(* IEC 61131-3 sources: codesys/project-view/Device/Plc Logic/Application/000-模组/本项目, 8 files *)

(* ---- FC_ArrayBoolHasTrue.st ---- *)
//布尔数组里面至少有一个值为true的话，函数返回TRUE
FUNCTION FC_ArrayBoolHasTrue : BOOL
VAR_IN_OUT
	abArray							: ARRAY[*] OF BOOL;
END_VAR

VAR
	i								: DINT;
END_VAR
// --- implementation ---
FOR i := LOWER_BOUND(abArray,1) TO UPPER_BOUND(abArray,1) DO
	IF abArray[i] THEN
		FC_ArrayBoolHasTrue := TRUE;
		RETURN;
	END_IF
END_FOR

FC_ArrayBoolHasTrue := FALSE;
END_FUNCTION

(* ---- FC_IsInArea.st ---- *)
FUNCTION FC_IsInArea : BOOL
VAR_INPUT
	LR_Pos							: REAL;//当前左右位置
	UD_Pos							: REAL;//当前上下位置

	LeftLimit						: REAL;//左边限位，LR_Pos要大于等于此变量
	RightLimit						: REAL;//右边限位，LR_Pos要小于等于此变量
	UpLimit							: REAL;//上边限位，UD_Pos要小于等于此变量
	DownLimit						: REAL;//下边限位，UD_Pos要大于等于此变量
END_VAR
VAR
END_VAR
// --- implementation ---
//判断是否在此平面范围内

IF (LeftLimit <= LR_Pos AND LR_Pos <= RightLimit) AND
	(DownLimit <= UD_Pos AND UD_Pos <= UpLimit) THEN

	FC_IsInArea := TRUE;
ELSE
	FC_IsInArea := FALSE;
END_IF
END_FUNCTION

(* ---- FC_StringConnect.st ---- *)
//输出 STRING = sStr1 + sStr2 + sStr3 + sStr4 +sStr5
FUNCTION FC_StringConnect : STRING
VAR_INPUT
	sStr1						: STRING:='';
	sStr2						: STRING:='';
	sStr3						: STRING:='';
	sStr4						: STRING:='';
	sStr5						: STRING:='';

END_VAR

VAR
	temp						: STRING;

END_VAR
// --- implementation ---
//temp := sStr1;

// StrConcatW(pstFrom:=ADR(wsContent_2) , pstTo:=ADR(temp) , iBufferSize:=TO_INT(SIZEOF(temp)) );
// StrConcatW(pstFrom:=ADR(wsContent_3) , pstTo:=ADR(temp) , iBufferSize:=TO_INT(SIZEOF(temp)) );

temp := CONCAT(STR1:=sStr1 , STR2:=sStr2 );
temp := CONCAT(STR1:=temp , STR2:=sStr3 );
temp := CONCAT(STR1:=temp , STR2:=sStr4 );
temp := CONCAT(STR1:=temp , STR2:=sStr5 );

FC_StringConnect := temp;
END_FUNCTION

(* ---- FC_WordToReal.st ---- *)
FUNCTION FC_WordToReal : REAL
VAR_INPUT
	arrRegisters0 : WORD;
	arrRegisters1 : WORD;
END_VAR
VAR
	dwCombined: DWORD;              // 合并后的DWORD
    rResult: REAL;                  // 输出浮点数
    pReal: POINTER TO REAL;         // 类型转换指针
    bIsBigEndian: BOOL := TRUE;     // 字节序配置开关
END_VAR
// --- implementation ---
// 寄存器合并与转换逻辑
IF bIsBigEndian THEN
    dwCombined := SHL(WORD_TO_DWORD(arrRegisters0), 16) OR arrRegisters1;
ELSE
    dwCombined := SHL(WORD_TO_DWORD(arrRegisters0), 16) OR arrRegisters1;
END_IF

pReal := ADR(dwCombined);           // 获取内存地址
FC_WordToReal := pReal^;                  // 指针解引用
END_FUNCTION

(* ---- FB_DelayInvert.st ---- *)
//X维持设定的初始值，直到指定时间结束，取反。
//若中途取消动作，X保持设定的初始值。
FUNCTION_BLOCK FB_DelayInvert
VAR_IN_OUT
	X							: BOOL;
END_VAR

VAR_INPUT
	bStart						: BOOL;
	bStop						: BOOL;

	bInitValue					: BOOL;//初始值
	tDelay						: TIME:=T#1S;

END_VAR

VAR_OUTPUT
END_VAR

VAR
	timer						: TON;
	R_TRIG_Start				: R_TRIG;
	R_TRIG_Stop					: R_TRIG;

END_VAR
// --- implementation ---
//定时器FB块
timer();

//启动
R_TRIG_Start(CLK:=bStart);
IF R_TRIG_Start.Q THEN
	X := bInitValue;
	timer.PT := tDelay;
	timer.IN := TRUE;
	bStart := FALSE;
END_IF

//定时器计时中（触发动作），中途取消动作，X维持初始值
R_TRIG_Stop(CLK:=bStop);
IF R_TRIG_Stop.Q AND timer.IN THEN
	X := bInitValue;
	timer.IN := FALSE;
END_IF

//时间到，取反
IF timer.Q THEN
	X := NOT X;
	timer.IN := FALSE;
END_IF
END_FUNCTION_BLOCK

(* ---- FB_Overtime.st ---- *)
FUNCTION_BLOCK FB_Overtime
VAR_INPUT
	bEnable						: BOOL;
	tTimeSet					: TIME:=T#1S;//定时时间
	iMode						: INT:=0;//超时后，0模式的bEnable变false，输出跟着变false；1模式的bEnable变false，输出不变，需要bReset复位。
	bReset						: BOOL;//上升沿将输出复位为false，仅1模式有效
END_VAR

VAR_OUTPUT
	bOvertime					: BOOL;
END_VAR

VAR
	tTimer						: TON;
	R_TRIG_1						: R_TRIG;
	R_TRIG_2						: R_TRIG;
END_VAR
// --- implementation ---
tTimer(IN:=bEnable , PT:= tTimeSet);
R_TRIG_1(CLK:=tTimer.Q);
R_TRIG_2(CLK:=bReset);

IF iMode = 0 THEN
	IF tTimer.Q THEN
		bOvertime:=TRUE;
	ELSE
		bOvertime:=FALSE;
	END_IF

ELSIF iMode = 1 THEN
	IF R_TRIG_1.Q THEN
		bOvertime:=TRUE;
	END_IF
	IF R_TRIG_2.Q THEN
		bOvertime:=false;
	END_IF

END_IF
END_FUNCTION_BLOCK

(* ---- FB_TcpClient_Free_1.st ---- *)
FUNCTION_BLOCK FB_TcpClient_Free_1
VAR_INPUT
	xConnect			:BOOL;				//连接
	xDisConnect			:BOOL;				//断开连接
	xReset				:BOOL;				//复位
	strIP				:STRING;			//IP
	uiPort				:UINT;				//端口号
	xSend				:BOOL;				//发送
	pbySendData			:POINTER TO BYTE;	//发送数据变量容器起始地址
	uxiSendDataSize		:__UXINT;			//发送数据变量容器大小
	uxiSendLenght		:__UXINT;			//发送数据长度
	pbyReceiveData		:POINTER TO BYTE;	//接收数据变量容器起始地址
	uxiReceiveDataSize	:__UXINT;			//接收数据变量容器大小
END_VAR
VAR_OUTPUT
	xBusy				:BOOL;				//运行中
	xConnected			:BOOL;				//已连接
	xError				:BOOL;				//错误
	xSendDone			:BOOL;				//发送完毕
	udiNumOfSend		:UDINT;				//发送次数（满4294967295自动清零）
	xReceiveDone		:BOOL;				//接收完毕
	udiNumOfReceive		:UDINT;				//接收次数（满4294967295自动清零）
	udiReceiveLenght	:UDINT;				//接收数据长度
END_VAR
VAR
	iStep			:INT;
	udiIndex		:UDINT;;
	fbClient		:TCP.Connector;
	eClientError	:TCP.ERROR;
	rtrigSend		:Standard.R_TRIG;
	eSendError		:TCP.ERROR;
	rtrigReceive	:Standard.R_TRIG;
	eReceiveError	:TCP.ERROR;
	xiReceiveLen	:__XINT;
	pby1			:POINTER TO BYTE;
	ton1:		Standard.TON;
END_VAR
// --- implementation ---
// ton1(IN:= TRUE, PT:= T#5000MS, Q=> , ET=> );
// IF NOT ton1.Q THEN
// 	RETURN;
// END_IF

IF xDisConnect THEN
	iStep:=0;
END_IF

//work step
CASE iStep OF

0:	//start
	fbClient.Disconnect();
	fbClient.Reset();
	RESET();
	xBusy:=FALSE;
	IF xConnect AND NOT xDisConnect THEN
		START();
		xBusy:=TRUE;
		iStep:=10;
	END_IF

10:	//wait connect
	eClientError:=fbClient.Connect(sIPAddress:= strIP, uiPort:= uiPort, pStream=> );
	IF eClientError = TCP.ERROR.NO_ERROR THEN
		xConnected:=TRUE;
		iStep:=20;
	ELSIF xReset THEN
		iStep:=0;
	END_IF

20:	//work
	RECEIVE();
	SEND();

30:	//error
	fbClient.Disconnect();
	fbClient.Reset();
	xConnected:=FALSE;
	xError:=TRUE;
	IF xReset THEN
		RESET();
		START();
		iStep:=10;
	END_IF

END_CASE
END_FUNCTION_BLOCK

ACTION SEND:
rtrigSend(CLK:= xSend, Q=> );
//没有触发send功能，把成功标志位置false
IF NOT xSend THEN
	xSendDone:=FALSE;
END_IF
IF rtrigSend.Q THEN
	//发送次数++1
	udiNumOfSend:=udiNumOfSend+1;
	IF udiNumOfSend=4294967295 THEN
		udiNumOfSend:=0;
	END_IF
	//判断发送长度，防止发送长度超越变量容器大小
	IF uxiSendLenght > uxiSendDataSize THEN
		eSendError:=fbClient._Stream.Send(pbyBuffer:= pbySendData, diBufferSize:= __UXINT_TO_DINT(uxiSendDataSize), diSent=> );
	ELSE
		eSendError:=fbClient._Stream.Send(pbyBuffer:= pbySendData, diBufferSize:= __UXINT_TO_DINT(uxiSendLenght), diSent=> );
	END_IF
	//判断发送结果
	IF eSendError = TCP.ERROR.NO_ERROR THEN
		xSendDone:=TRUE;
	ELSE
		iStep:=30;
	END_IF
END_IF
END_ACTION

ACTION RECEIVE:
//启动receive功能
eReceiveError:=fbClient._Stream.Receive(pbyBuffer:= pbyReceiveData, diBufferSize:= __UXINT_TO_DINT(uxiReceiveDataSize), diReceived=> xiReceiveLen);
rtrigReceive(CLK:= eReceiveError=TCP.ERROR.NO_ERROR , Q=> );
IF rtrigReceive.Q THEN
	//发送次数++1
	udiNumOfReceive:=udiNumOfReceive+1;
	IF udiNumOfReceive=4294967295 THEN
		udiNumOfReceive:=0;
	END_IF
	//触发接收标志位时，对接收数据操作。把不属于本次接收数据长度以外的数据清除
	FOR udiIndex:=__XINT_TO_UDINT(xiReceiveLen) TO (__UXINT_TO_UDINT(uxiReceiveDataSize)-1) BY 1 DO
		pby1:=pbyReceiveData+udiIndex;
		pby1^:=0;
	END_FOR
	//输出接收数据长度
	udiReceiveLenght:=__XINT_TO_UDINT(xiReceiveLen);
END_IF
//输出接收成功标志位，上升沿
xReceiveDone:=rtrigReceive.Q;
//receive功能错误判定
IF eReceiveError <> TCP.ERROR.NO_ERROR AND eReceiveError <> TCP.ERROR.PENDING THEN
	iStep:=30;
END_IF
END_ACTION

ACTION RESET:
//复位各类标志位
xConnected:=FALSE;
xError:=FALSE;
xSendDone:=FALSE;
xReceiveDone:=FALSE;
udiReceiveLenght:=0;
udiNumOfSend:=0;
udiNumOfReceive:=0;

//复位功能rtrig
rtrigReceive(CLK:= FALSE, Q=> );
rtrigSend(CLK:= FALSE, Q=> );

//复位功能fun状态
eClientError:=TCP.ERROR.NO_ERROR;
eReceiveError:=TCP.ERROR.NO_ERROR;
eSendError:=TCP.ERROR.NO_ERROR;
END_ACTION

ACTION START:
//启动前，会对 发送与接收 容器进行清除数据
FOR udiIndex:=0 TO (__UXINT_TO_UDINT(uxiSendDataSize)-1) BY 1 DO
	pby1:=pbySendData+udiIndex;
	pby1^:=0;
END_FOR
FOR udiIndex:=0 TO (__UXINT_TO_UDINT(uxiReceiveDataSize)-1) BY 1 DO
	pby1:=pbyReceiveData+udiIndex;
	pby1^:=0;
END_FOR
END_ACTION

(* ---- FB_ValueChanged.st ---- *)
//监控变量的值是否发生改变
FUNCTION_BLOCK FB_ValueChanged
VAR_INPUT
	pValue						: POINTER TO BYTE;
	uxiSize						: __UXINT;
END_VAR

VAR_OUTPUT
	bHasChanged					: BOOL;//变量值发生改变，该输出变量保持一个周期 true
END_VAR

VAR
	bFirstScan					: BOOL;
	pOrigin						: POINTER TO BYTE;//记录变量上一个周期的值

END_VAR
// --- implementation ---
//初次上电，分配与 pValue 相同长度的内存
IF NOT bFirstScan THEN
	pOrigin := SM3_Basic.SysMemAllocData(szComponent:='pOrigin' , udiSize:=uxiSize , pResult:=0 );
	bFirstScan := TRUE;
END_IF

//比较内存值
IF 0 <> SM3_Basic.SysMemCmp(pBuffer1:=pOrigin , pBuffer2:=pValue , udiCount:=uxiSize ) THEN
	SM3_Basic.SysMemCpy(pDest:=pOrigin , pSrc:=pValue , udiCount:=uxiSize );//从指针层面，将新值复制到pOrigin
	bHasChanged := TRUE;
ELSE
	bHasChanged := FALSE;
END_IF
END_FUNCTION_BLOCK
